(* IEC 61131-3 sources: plc-iiot-stack/src/POUs/Iiot/F_IiotCmdKind, 2 files *)

(* ---- F_IiotCmdKind.decl.st ---- *)
// Назначение: вид команды по полю value: значение (SpeedSp, SubstValue), маска (AckReq,
//             ShelveReq, UnshelveReq) или импульс (остальные).
// Автор:      kr0nsch
// Версия:     0.1.0
// Документ:   docs/plc_mqtt.md, раздел «Команды»
FUNCTION F_IiotCmdKind : E_IiotCmdKind
VAR_INPUT
    eCommand : E_IiotCommand;
END_VAR

(* ---- F_IiotCmdKind.impl.st ---- *)
CASE eCommand OF
    E_IiotCommand.SpeedSp, E_IiotCommand.SubstValue:
        F_IiotCmdKind := E_IiotCmdKind.Value;
    E_IiotCommand.AckReq, E_IiotCommand.ShelveReq, E_IiotCommand.UnshelveReq:
        F_IiotCmdKind := E_IiotCmdKind.Mask;
ELSE
    F_IiotCmdKind := E_IiotCmdKind.Pulse;
END_CASE
